(* IEC 61131-3 sources: repolevel_ST_code_completion/output/0127完整版本_带planner/repoeval_electronic_gear_motion/readful_result_before_fix, 3 files *)

(* ---- FB_DualAxisPower.st ---- *)
FUNCTION_BLOCK FB_DualAxisPower
VAR_INPUT
	Axis1			:	AXIS_REF;		//轴1引用
	Axis2			:	AXIS_REF;		//轴2引用
	bEnable			:	BOOL := TRUE;	//使能信号
END_VAR
VAR_OUTPUT
	bAxis1Ready		:	BOOL;			//轴1准备就绪
	bAxis2Ready		:	BOOL;			//轴2准备就绪
	bBothReady		:	BOOL;			//两轴都准备就绪
	bError			:	BOOL;			//错误标志
END_VAR
VAR
	fbPower1		:	MC_Power;		//轴1电源控制
	fbPower2		:	MC_Power;		//轴2电源控制
END_VAR

IF NOT bEnable THEN
	bAxis1Ready := FALSE;
	bAxis2Ready := FALSE;
	bBothReady := FALSE;
	bError := FALSE;
	RETURN;
END_IF

// 执行轴1电源控制
fbPower1(
	Axis := Axis1,
	Enable := bEnable,
	bDriveStart := TRUE,
	bRegulatorOn := TRUE
);

// 执行轴2电源控制
fbPower2(
	Axis := Axis2,
	Enable := bEnable,
	bDriveStart := TRUE,
	bRegulatorOn := TRUE
);

// 检查轴1状态
IF NOT fbPower1.Status OR fbPower1.Error THEN
	bAxis1Ready := FALSE;
	bError := TRUE;
	RETURN;
ELSE
	bAxis1Ready := TRUE;
END_IF

// 检查轴2状态
IF NOT fbPower2.Status OR fbPower2.Error THEN
	bAxis2Ready := FALSE;
	bError := TRUE;
	RETURN;
ELSE
	bAxis2Ready := TRUE;
END_IF

// 更新两轴准备状态
bBothReady := bAxis1Ready AND bAxis2Ready;

// 检查最终状态
IF bBothReady AND NOT bError THEN
	RETURN;
END_IF
END_FUNCTION_BLOCK

(* ---- FB_GearCoupling.st ---- *)
FUNCTION_BLOCK FB_GearCoupling
VAR_INPUT
	Master				:	AXIS_REF;		//主轴引用
	Slave				:	AXIS_REF;		//从轴引用
	bCouple				:	BOOL;			//TRUE=耦合，FALSE=解耦
	nRatioNumerator		:	INT := 1;		//传动比分子
	nRatioDenominator	:	INT := 1;		//传动比分母
	rAcceleration		:	REAL := 10000.0;//加速度
	rDeceleration		:	REAL := 10000.0;//减速度
END_VAR
VAR_OUTPUT
	bInGear				:	BOOL;			//耦合状态
	bCouplingDone		:	BOOL;			//耦合完成
	bDecouplingDone		:	BOOL;			//解耦完成
	bError				:	BOOL;			//错误标志
	nErrorID			:	DWORD;			//错误代码
END_VAR
VAR
	fbGearIn			:	MC_GearIn;		//齿轮耦合功能块
	fbGearOut			:	MC_GearOut;		//齿轮解耦功能块
	bLastCouple			:	BOOL;			//上次耦合状态
	bCoupleRising		:	BOOL;			//耦合上升沿
	bCoupleFalling		:	BOOL;			//耦合下降沿
END_VAR

// 检测耦合信号的边沿
bCoupleRising := bCouple AND NOT bLastCouple;
bCoupleFalling := NOT bCouple AND bLastCouple;
bLastCouple := bCouple;

// 耦合逻辑
IF bCouple THEN
	IF bCoupleRising THEN
		// 配置齿轮耦合功能块
		fbGearIn.Master := Master;
		fbGearIn.Slave := Slave;
		fbGearIn.RatioNumerator := nRatioNumerator;
		fbGearIn.RatioDenominator := nRatioDenominator;
		fbGearIn.Acceleration := rAcceleration;
		fbGearIn.Deceleration := rDeceleration;
		fbGearIn.Execute := TRUE;
	END_IF

	// 检查耦合状态
	IF fbGearIn.Done THEN
		bInGear := TRUE;
		bCouplingDone := TRUE;
		bError := FALSE;
		nErrorID := 0;
	ELSIF fbGearIn.Error THEN
		bError := TRUE;
		nErrorID := fbGearIn.ErrorID;
	END_IF
ELSE
	// 解耦逻辑
	IF bCoupleFalling THEN
		// 配置齿轮解耦功能块
		fbGearOut.Master := Master;
		fbGearOut.Slave := Slave;
		fbGearOut.Execute := TRUE;
	END_IF

	// 检查解耦状态
	IF fbGearOut.Done THEN
		bInGear := FALSE;
		bDecouplingDone := TRUE;
		bError := FALSE;
		nErrorID := 0;
	ELSIF fbGearOut.Error THEN
		bError := TRUE;
		nErrorID := fbGearOut.ErrorID;
	END_IF
END_IF
END_FUNCTION_BLOCK

(* ---- FB_GearMotionControl.st ---- *)
FUNCTION_BLOCK FB_GearMotionControl
VAR_INPUT
	MasterAxis			:	AXIS_REF;		//主轴引用
	SlaveAxis			:	AXIS_REF;		//从轴引用
	bStart				:	BOOL;			//启动信号
	bStop				:	BOOL;			//停止信号
	nRatioNumerator		:	INT := 1;		//传动比分子
	nRatioDenominator	:	INT := 1;		//传动比分母
	nDirection			:	INT := 1;		//运动方向（1=正向，-1=反向）
	rVelocity			:	REAL := 360.0;	//主轴速度
	rAcceleration		:	REAL := 10000.0;//加速度
	rDeceleration		:	REAL := 10000.0;//减速度
END_VAR
VAR_OUTPUT
	bRunning			:	BOOL;			//运行中
	bReady				:	BOOL;			//准备就绪（可以启动）
	bError				:	BOOL;			//错误标志
	nCurrentState		:	BYTE;			//当前状态
END_VAR
VAR
	fbPowerMgr			:	FB_DualAxisPower;	//双轴电源管理
	fbGearCtrl			:	FB_GearCoupling;	//齿轮耦合控制
	fbMoveVel			:	MC_MoveVelocity;	//速度运动
	fbHaltMaster		:	MC_Halt;			//主轴停止
	fbHaltSlave			:	MC_Halt;			//从轴停止
	fbStartRtrig		:	R_TRIG;				//启动上升沿
	fbStopRtrig			:	R_TRIG;				//停止上升沿
	nState				:	BYTE;				//内部状态机
	rSlaveVelocity		:	REAL;				//从轴速度
END_VAR

fbStartRtrig(CLK := bStart);
fbStopRtrig(CLK := bStop);

IF fbStopRtrig.Q THEN
	// 停止信号优先处理
	fbHaltMaster(Execute := TRUE, Axis := MasterAxis, Deceleration := rDeceleration);
	fbHaltSlave(Execute := TRUE, Axis := SlaveAxis, Deceleration := rDeceleration);
	bRunning := FALSE;
	bReady := FALSE;
	nState := 0;
	RETURN;
END_IF

IF fbStartRtrig.Q THEN
	// 检查输入参数合法性
	IF nRatioNumerator = 0 OR nRatioDenominator = 0 OR (nDirection <> 1 AND nDirection <> -1) THEN
		bError := TRUE;
		RETURN;
	END_IF;

	// 计算从轴速度
	rSlaveVelocity := rVelocity * nRatioNumerator / nRatioDenominator * nDirection;

	// 设置主轴和从轴运动参数
	fbMoveVel(Execute := TRUE, Axis := MasterAxis, Velocity := rVelocity, Acceleration := rAcceleration, Deceleration := rDeceleration);
	fbGearCtrl(Execute := TRUE, Master := MasterAxis, Slave := SlaveAxis, RatioNumerator := nRatioNumerator, RatioDenominator := nRatioDenominator);

	// 更新状态
	bRunning := TRUE;
	bReady := FALSE;
	nState := 1;
	RETURN;
END_IF;

CASE nState OF
	0: // 等待轴准备就绪
		IF fbPowerMgr.Axis1Ready AND fbPowerMgr.Axis2Ready THEN
			bReady := TRUE;
		END_IF;

	1: // 运行中
		IF NOT fbMoveVel.Busy THEN
			bRunning := FALSE;
			bReady := TRUE;
			nState := 0;
		END_IF;

		IF fbMoveVel.Error OR fbGearCtrl.Error THEN
			bError := TRUE;
			fbHaltMaster(Execute := TRUE, Axis := MasterAxis, Deceleration := rDeceleration);
			fbHaltSlave(Execute := TRUE, Axis := SlaveAxis, Deceleration := rDeceleration);
			nState := 0;
		END_IF;
END_CASE;
END_FUNCTION_BLOCK
